// TIA Portal project "EXO" (V16)

(* hardware
DEVICE "Station S7300/ET200M_1"  S7-300 station
   slot 0: "Châssis_0"  Rail  6ES7 390-1***0-0AA0
   slot 2: "PLC_1"  CPU 314C-2 PN/DP  6ES7 314-6EH04-0AB0  V3.3
      slot 2: "Interface PROFINET_1"  PN-IO
         slot 1: "Port_1"  Port
         slot 2: "Port_2"  Port
      slot 5: "DI 24/DO 16_1"  DI24/DO16
      slot 6: "AI 5/AO 2_1"  AI5/AO2
      slot 7: "Comptage_1"  Counter
      slot 8: "Positionnement_1"  Positioning
*)

// ===== PLC "PLC_1"  CPU 314C-2 PN/DP =====

VAR_GLOBAL   // PLC tag table "Table de variables standard"
   "START" AT %I0.0 : Bool;
   "BP_stop" AT %I0.1 : Bool;
   "BP_reset" AT %I0.2 : Bool;
   "H1" AT %Q0.1 : Bool;
   "MOTEUR" AT %Q0.2 : Bool;
   "M" AT %M0.1 : Bool;
END_VAR

ORGANIZATION_BLOCK "Main"   // OB1, LAD
TITLE = "Main Program Sweep (Cycle)"
{ S7_Optimized_Access := 'FALSE' }
VERSION : 0.1
   VAR_TEMP
      OB1_EV_CLASS : Byte;   // Bits 0-3 = 1 (Coming event), Bits 4-7 = 1 (Event class 1)
      OB1_SCAN_1 : Byte;   // 1 (Cold restart scan 1 of OB 1), 3 (Scan 2-n of OB 1)
      OB1_PRIORITY : Byte;   // Priority of OB Execution
      OB1_OB_NUMBR : Byte;   // 1 (Organization block 1, OB1)
      OB1_RESERVED_1 : Byte;   // Reserved for system
      OB1_RESERVED_2 : Byte;   // Reserved for system
      OB1_PREV_CYCLE : Int;   // Cycle time of previous OB1 scan (milliseconds)
      OB1_MIN_CYCLE : Int;   // Minimum cycle time of OB1 (milliseconds)
      OB1_MAX_CYCLE : Int;   // Maximum cycle time of OB1 (milliseconds)
      OB1_DATE_TIME : Date_And_Time;   // Date and time OB1 started
   END_VAR
BEGIN

REGION Network 1
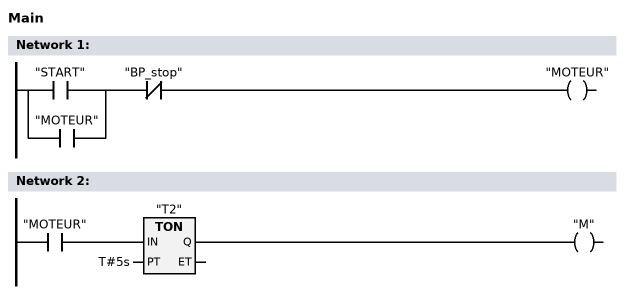
   RUNG wire#powerrail
      Contact( "START" )
      wire#w1
      I_Contact( "BP_stop" )
      Coil( "MOTEUR" )
   END_RUNG
   RUNG wire#powerrail
      Contact( "MOTEUR" )
   END_RUNG wire#w1
   // the same network as SCL:
   "MOTEUR" := ("START" OR "MOTEUR") AND NOT "BP_stop";
END_REGION

REGION Network 2
   "T2".TON(IN := "MOTEUR", PT := T#5s);
   "M" := "T2".Q;
END_REGION
END_ORGANIZATION_BLOCK